(* IEC 61131-3 sources: PLC-Programming-using-OpenPLC/01.Start/build, 1 file *)

(* ---- generated_plc.st ---- *)
PROGRAM program0
  VAR
    X100 : BOOL;
    Y100 : BOOL;
  END_VAR

  Y100 := X100;
END_PROGRAM

CONFIGURATION Config0

  RESOURCE Res0 ON PLC
    TASK task0(INTERVAL := T#20ms,PRIORITY := 0);
    PROGRAM instance0 WITH task0 : program0;
  END_RESOURCE
END_CONFIGURATION
